SUBAPPLICATION AX_TO_QXA_BG_PUBLISH_OPT (* Wie AX_TO_QXA_BG_PUBLISH, aber physischer Ausgang getrennt gegatet: Hintergrund+State-Publish laufen immer (QI/INIT), nur DigitalOutput haengt an QI_Output/INIT_Output (z.B. Option Klassisch vs. PVEA auf gemeinsamem Pin). *)
  (* Standard: 61499-2; Description: Copyright (c) 2026 Meisterschulen am Ostbahnhof This program and the accompanying materials are made available under the terms of the Eclipse Public License 2.0 which is available at https://www.eclipse.org/legal/epl-2.0/ SPDX-License-Identifier: EPL-2.0 *)
  (* Version 1.0, 2026-10-16, Franz Höpfinger, Meisterschulen am Ostbahnhof, Kopie von AX_TO_QXA_BG_PUBLISH v1.2 (Franz: 'Die Lib Typen KOPIEREN und die Kopie aendern') - QI/INIT gelten nur noch fuer Hintergrund+Publish, neuer QI_Output/INIT_Output/INITO_Output/QO_Output nur fuer DigitalOutput. Grund: bei Igel/Elevator=PVEA blieb mit dem Ausgang auch SoftKey-Hintergrund und State-Publish tot. *)
  PACKAGE MyLib::sys;
  IMPORT isobus::UT::Q::const::IDs::ID_NULL;
  IMPORT logiBUS::io::DQ::logiBUS_DO;
  IMPORT logiBUS::io::DQ::logiBUS_DO_S;
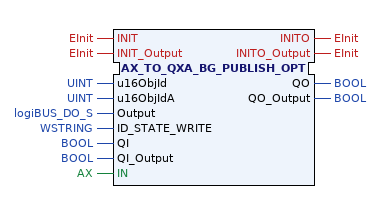
  EVENT_INPUT
    INIT : EInit; (* Initialisierung Hintergrund+Publish (Anzeige) - typisch sofort beim Boot *)
    INIT_Output : EInit; (* Initialisierung physischer Ausgang - typisch von der Option getrieben *)
  END_EVENT
  EVENT_OUTPUT
    INITO : EInit; (* Anzeige initialisiert - echtes Confirm von PUBLISH_STATE.INITO *)
    INITO_Output : EInit; (* Ausgang initialisiert - echtes Confirm von DigitalOutput.INITO *)
  END_EVENT
  VAR_INPUT
    u16ObjId : UINT := ID_NULL; (* Object ID Softkey - traegt die Hintergrundfarbe *)
    u16ObjIdA : UINT := ID_NULL; (* Object ID AuxFunction2 (Joystick) - zeigt Hintergrundfarbe am Aux-Handle mit *)
    Output : logiBUS::io::DQ::logiBUS_DO_S := logiBUS_DO::Invalid; (* Identify the Output Output_Q1..Q12 *)
    ID_STATE_WRITE : WSTRING; (* Lokale Publish-Adresse (ACTION=WRITE) fuer den Zustand - wird von Web-Client/Dashboard remote abonniert *)
    QI : BOOL := TRUE; (* Qualifier Hintergrund+Publish (Anzeige) *)
    QI_Output : BOOL := TRUE; (* Qualifier nur fuer den physischen Ausgang - FALSE gibt den Pin frei *)
  END_VAR
  VAR_OUTPUT
    QO : BOOL; (* Quality Output Anzeige (AND aus GreenWhiteBackground_AX/PUBLISH_STATE) *)
    QO_Output : BOOL; (* Quality Output physischer Ausgang (DigitalOutput.QO) *)
  END_VAR
  SOCKETS
    IN : adapter::types::unidirectional::AX; (* Fertiger AX-Zustand - wird auf Ausgang+Hintergrund+Publish verteilt *)
  END_SOCKETS
  FBS
    AX_SPLIT_3 : adapter::events::unidirectional::AX_SPLIT_3;
    DigitalOutput : logiBUS::io::DQ::logiBUS_QXA;
    PUBLISH_STATE : adapter::net::AX_PUBLISH_1;
    AND_QO : iec61131::booleanOperators::AND_BOOL_2;
  END_FBS
  SUBAPPS
    GreenWhiteBackground_AX : MyLib::sys::GreenWhiteBackground3_AX;
  END_SUBAPPS
  EVENT_CONNECTIONS
    INIT_Output TO DigitalOutput.INIT;
    DigitalOutput.INITO TO INITO_Output;
    INIT TO GreenWhiteBackground_AX.INIT;
    GreenWhiteBackground_AX.INITO TO PUBLISH_STATE.INIT;
    PUBLISH_STATE.INITO TO INITO;
    PUBLISH_STATE.INITO TO AND_QO.REQ;
  END_CONNECTIONS
  DATA_CONNECTIONS
    u16ObjId TO GreenWhiteBackground_AX.u16ObjId;
    u16ObjIdA TO GreenWhiteBackground_AX.u16ObjIdA;
    Output TO DigitalOutput.Output;
    ID_STATE_WRITE TO PUBLISH_STATE.ID;
    QI_Output TO DigitalOutput.QI;
    QI TO PUBLISH_STATE.QI;
    QI TO GreenWhiteBackground_AX.QI;
    GreenWhiteBackground_AX.QO TO AND_QO.IN1;
    PUBLISH_STATE.QO TO AND_QO.IN2;
    AND_QO.OUT TO QO;
    DigitalOutput.QO TO QO_Output;
  END_CONNECTIONS
  ADAPTER_CONNECTIONS
    IN TO AX_SPLIT_3.IN;
    AX_SPLIT_3.OUT1 TO DigitalOutput.OUT;
    AX_SPLIT_3.OUT2 TO GreenWhiteBackground_AX.DI1;
    AX_SPLIT_3.OUT3 TO PUBLISH_STATE.IN;
  END_CONNECTIONS
END_SUBAPPLICATION
